Fanuc KAREL source: KA00138.KL

PROGRAM KA00138
%NOLOCKGROUP
VAR
  SRC: ARRAY[2] OF SHORT
  DST: XYZWPR
BEGIN
  SRC[1] = 2
  DST = SRC[1]
END KA00138
